(* IEC 61131-3 sources: SRCI_CLIENT_PLC/RobotLibrary/Library/POUs/Calculation/MC_LoadMeasurementSequential/Structures, 4 files *)

(* ---- LoadMeasurementSequentialOutCmd.st ---- *)
{attribute 'pack_mode' := '1'}
// -------------------------------------------------------------------------
//  SRCI Robot Library
// -------------------------------------------------------------------------
//
//  Object:      LoadMeasurementSequentialOutCmd
//  Author:      Thorsten Brach
//  Date:        2024-06-20
//
//  Description:
//
//
//  Copyright:
//    (C) 2024 Thorsten Brach. All rights reserved
//             Licensed under the MIT License.
//
//  Disclaimer:
//    This project is provided without any guarantee and can be used for
//    private and commercial purposes. Any use is at the user’s
//    own risk and responsibility.
//
// -------------------------------------------------------------------------
TYPE LoadMeasurementSequentialOutCmd :
STRUCT
  /// FB is returning a unique ID for the cal led measurement.
  MeasuringID        : UINT;
  /// Measured load data (see chapter 5.5.6.4)
  LoadData           : LoadData;
  /// Load data available
  LoadDataAvailable : BOOL;
END_STRUCT
END_TYPE

(* ---- LoadMeasurementSequentialParCmd.st ---- *)
{attribute 'pack_mode' := '1'}
// -------------------------------------------------------------------------
//  SRCI Robot Library
// -------------------------------------------------------------------------
//
//  Object:      LoadMeasurementSequentialParCmd
//  Author:      Thorsten Brach
//  Date:        2024-06-20
//
//  Description:
//
//
//  Copyright:
//    (C) 2024 Thorsten Brach. All rights reserved
//             Licensed under the MIT License.
//
//  Disclaimer:
//    This project is provided without any guarantee and can be used for
//    private and commercial purposes. Any use is at the user’s
//    own risk and responsibility.
//
// -------------------------------------------------------------------------
TYPE LoadMeasurementSequentialParCmd :
STRUCT
  /// Define which step of the load estimation should be executed:
  Mode               : LoadMeasurementSteps;
  /// Define which mass is expected as a result of the load measurement
  Mass               : REAL;
END_STRUCT
END_TYPE

(* ---- LoadMeasurementSequentialRecvData.st ---- *)
{attribute 'pack_mode' := '1'}
// -------------------------------------------------------------------------
//  SRCI Robot Library
// -------------------------------------------------------------------------
//
//  Object:      LoadMeasurementSequentialRecvData
//  Author:      Thorsten Brach
//  Date:        2024-06-20
//
//  Description:
//
//
//  Copyright:
//    (C) 2024 Thorsten Brach. All rights reserved
//             Licensed under the MIT License.
//
//  Disclaimer:
//    This project is provided without any guarantee and can be used for
//    private and commercial purposes. Any use is at the user’s
//    own risk and responsibility.
//
// -------------------------------------------------------------------------
TYPE LoadMeasurementSequentialRecvData EXTENDS RspHeader :
STRUCT
  /// FB is returning a unique ID for the cal led measurement.
  MeasuringID       : UINT;
  /// Measured load data (see chapter 5.5.6.4)
  LoadData          : LoadData;
  /// Load data available
  LoadDataAvailable : BOOL;
END_STRUCT
END_TYPE

(* ---- LoadMeasurementSequentialSendData.st ---- *)
{attribute 'pack_mode' := '1'}
// -------------------------------------------------------------------------
//  SRCI Robot Library
// -------------------------------------------------------------------------
//
//  Object:      LoadMeasurementSequentialSendData
//  Author:      Thorsten Brach
//  Date:        2024-06-20
//
//  Description:
//
//
//  Copyright:
//    (C) 2024 Thorsten Brach. All rights reserved
//             Licensed under the MIT License.
//
//  Disclaimer:
//    This project is provided without any guarantee and can be used for
//    private and commercial purposes. Any use is at the user’s
//    own risk and responsibility.
//
// -------------------------------------------------------------------------
TYPE LoadMeasurementSequentialSendData EXTENDS CmdHeader:
STRUCT
    /// Define which mass is expected as a result of the load measurement
  Mass               : REAL;
  /// Define which step of the load estimation should be executed:
  Mode               : LoadMeasurementSteps;
END_STRUCT
END_TYPE
